TYPE ST_Mover :
STRUCT
	nId: DINT;
	nPhysicalId: DINT;
	nLoadBearing: DINT;
	nLength: DINT;
	nWidth: DINT;
	nClampLength: DINT;
	nClampwidth: DINT;
	nOffset: DINT;
	nMoverTolerance: DINT;
	nGap: DINT;
	nInitialPosition: DINT;
	nInitialRoad: DINT;
END_STRUCT
END_TYPE

(* stored: Version 1.1.0.1, ProductVersion 3.1.4024.12
   DUT ST_Mover: Id {7210eb91-4eb3-4d20-b2f0-8759a8a87dd5} *)
